(*
	One timed operation in a trace. Unlike a log record, a span has a lifecycle:
	  building - FB_Tracer owns it while the fluent chain fills it in,
	  running  - build hands it to the caller, who owns it while the work runs,
	  ended    - FB_Tracer.endSpan hands it to the provider for processing.
	The span owns every pointer member and releases them in free. A running span is read and
	changed only through FB_Tracer, such as getSpanContext, setSpanStatusOk and discardSpan,
	so callers never dereference it themselves. The methods left here belong to the tracing
	pipeline: the provider, samplers and processors.
*)
{attribute 'enable_dynamic_creation'}
FUNCTION_BLOCK FB_Span
VAR_INPUT
	// written by the tracer while the span is built
	name: POINTER TO FB_String;
	kind: E_SpanKind;
	startTimestamp: ULINT;
	endTimestamp: ULINT;
	traceId: POINTER TO FB_TraceId;
	spanId: POINTER TO FB_SpanId;
	traceState: POINTER TO FB_TraceState;

	// required if child span, must be omitted if root span
	parentSpanId: POINTER TO FB_SpanId;

	// describes the parent's remoteness, not this span's; see E_SpanFlags
	flags: UDINT;
	status: POINTER TO FB_Status;
END_VAR
VAR_OUTPUT
	attributes: FB_Attributes(maxCount := TcOtlp_GVL.DEFAULT_MAX_ATTRIBUTE_COUNT);
	links: FB_Links(maxCount := TcOtlp_GVL.DEFAULT_MAX_LINK_COUNT);
	resource: FB_Resource('');
	scope: FB_InstrumentationScope('', '', '');

	// span events have been deprecated, instead logs should be emitted with span context for correlation
	// events
	// droppedEventCount
END_VAR

(*
	Releases this span and clears the caller's pointer to it: call it as p^.delete(pSelf:=p).
	pSelf is cleared before the span is freed, so the caller never keeps a dangling pointer.
	A pointer to any other object is refused and left untouched, and nothing is released.
*)
METHOD delete : BOOL
VAR_IN_OUT
	pSelf: POINTER TO FB_Span;
END_VAR
VAR
	_pThis: POINTER TO FB_Span;
END_VAR
_pThis := THIS;
IF pSelf <> _pThis THEN
	RETURN;
END_IF

pSelf := 0;
__DELETE(_pThis);
delete := TRUE;
END_METHOD

//FB_Exit must be implemented explicitly. If there is an implementation, then the
//method is called before the controller removes the code of the function block instance
//(implicit call). The return value is not evaluated.
METHOD FB_Exit: BOOL
VAR_INPUT
    bInCopyCode: BOOL;  // TRUE: the exit method is called in order to leave the instance which will be copied afterwards (online change).
END_VAR
IF NOT bInCopyCode THEN
	THIS^.free();
END_IF
END_METHOD

(* Releases everything the span owns. Safe to call more than once. *)
METHOD free
IF THIS^.name <> 0 THEN THIS^.name^.delete(pSelf:=THIS^.name); END_IF
IF THIS^.traceId <> 0 THEN THIS^.traceId^.delete(pSelf:=THIS^.traceId); END_IF
IF THIS^.spanId <> 0 THEN THIS^.spanId^.delete(pSelf:=THIS^.spanId); END_IF
IF THIS^.traceState <> 0 THEN THIS^.traceState^.delete(pSelf:=THIS^.traceState); END_IF
IF THIS^.parentSpanId <> 0 THEN THIS^.parentSpanId^.delete(pSelf:=THIS^.parentSpanId); END_IF
IF THIS^.status <> 0 THEN THIS^.status^.delete(pSelf:=THIS^.status); END_IF
THIS^.attributes.free();
THIS^.links.free();
THIS^.scope.free();
THIS^.resource.free();
END_METHOD

(*
	Allocates a deep copy of this span, for a processor that keeps an ended span past onEnd.
	The copy owns copies of every member, so it stays valid after this span is released. This
	span is only read, apart from its links cursor. The caller owns pDest, which must be 0; on
	failure nothing is allocated and pDest is left alone.
*)
METHOD cloneTo : BOOL
VAR_IN_OUT
	pDest: POINTER TO FB_Span;
END_VAR
VAR_OUTPUT
	failureReason: E_SpanCloneFailureReason;
END_VAR
VAR
	_pClone: POINTER TO FB_Span;
	_pMessage: POINTER TO FB_String;
	_copied: BOOL;
	_attributesFailureReason: E_AttributesFailureReason;
	_linkFailureReason: E_LinkFailureReason;
END_VAR
cloneTo := FALSE;
failureReason := E_SpanCloneFailureReason.NA;

IF pDest <> 0 THEN
	failureReason := E_SpanCloneFailureReason.DESTINATION_ALREADY_ASSIGNED;
	RETURN;
END_IF

_pClone := __NEW(FB_Span);
IF _pClone = 0 THEN
	failureReason := E_SpanCloneFailureReason.MEMORY_ALLOCATION_FAILURE;
	RETURN;
END_IF

// the clone owns its members from here, so deleting it releases whatever was copied
_pClone^.kind := THIS^.kind;
_pClone^.startTimestamp := THIS^.startTimestamp;
_pClone^.endTimestamp := THIS^.endTimestamp;
_pClone^.flags := THIS^.flags;

_copied := (THIS^.name = 0 OR_ELSE ValueFactory.cloneString(
		pDest:=_pClone^.name,
		pSrc:=THIS^.name))
	AND_THEN (THIS^.traceId = 0 OR_ELSE ValueFactory.createTraceId(
		pDest:=_pClone^.traceId,
		pBytes:=ADR(THIS^.traceId^.bytes),
		nSize:=SIZEOF(THIS^.traceId^.bytes)))
	AND_THEN (THIS^.spanId = 0 OR_ELSE ValueFactory.createSpanId(
		pDest:=_pClone^.spanId,
		pBytes:=ADR(THIS^.spanId^.bytes),
		nSize:=SIZEOF(THIS^.spanId^.bytes)))
	AND_THEN (THIS^.parentSpanId = 0 OR_ELSE ValueFactory.createSpanId(
		pDest:=_pClone^.parentSpanId,
		pBytes:=ADR(THIS^.parentSpanId^.bytes),
		nSize:=SIZEOF(THIS^.parentSpanId^.bytes)))
	AND_THEN (THIS^.traceState = 0 OR_ELSE TraceStateFactory.clone(
		pDest:=_pClone^.traceState,
		pSrc:=THIS^.traceState))
	AND_THEN (THIS^.status = 0 OR_ELSE THIS^.status^.message = 0 OR_ELSE ValueFactory.cloneString(
		pDest:=_pMessage,
		pSrc:=THIS^.status^.message));
IF NOT _copied THEN
	IF _pMessage <> 0 THEN _pMessage^.delete(pSelf:=_pMessage); END_IF
	_pClone^.delete(pSelf:=_pClone);
	failureReason := E_SpanCloneFailureReason.VALUE_COPY_FAILURE;
	RETURN;
END_IF

IF THIS^.status <> 0 THEN
	_pClone^.status := __NEW(FB_Status(code:=THIS^.status^.code, message:=_pMessage));
	IF _pClone^.status = 0 THEN
		IF _pMessage <> 0 THEN _pMessage^.delete(pSelf:=_pMessage); END_IF
		_pClone^.delete(pSelf:=_pClone);
		failureReason := E_SpanCloneFailureReason.MEMORY_ALLOCATION_FAILURE;
		RETURN;
	END_IF
	_pMessage := 0;  // moved into the status
END_IF

IF NOT _pClone^.attributes.copyFrom(src:=THIS^.attributes, failureReason=>_attributesFailureReason) THEN
	_pClone^.delete(pSelf:=_pClone);
	IF _attributesFailureReason = E_AttributesFailureReason.MEMORY_ALLOCATION_FAILURE THEN
		failureReason := E_SpanCloneFailureReason.MEMORY_ALLOCATION_FAILURE;
	ELSE
		failureReason := E_SpanCloneFailureReason.ATTRIBUTE_COPY_FAILURE;
	END_IF
	RETURN;
END_IF

IF NOT _pClone^.links.copyFrom(src:=THIS^.links, failureReason=>_linkFailureReason) THEN
	_pClone^.delete(pSelf:=_pClone);
	IF _linkFailureReason = E_LinkFailureReason.MEMORY_ALLOCATION_FAILURE THEN
		failureReason := E_SpanCloneFailureReason.MEMORY_ALLOCATION_FAILURE;
	ELSE
		failureReason := E_SpanCloneFailureReason.LINK_COPY_FAILURE;
	END_IF
	RETURN;
END_IF

IF NOT _pClone^.resource.copyFrom(src:=THIS^.resource, failureResult=>_attributesFailureReason) THEN
	_pClone^.delete(pSelf:=_pClone);
	IF _attributesFailureReason = E_AttributesFailureReason.MEMORY_ALLOCATION_FAILURE THEN
		failureReason := E_SpanCloneFailureReason.MEMORY_ALLOCATION_FAILURE;
	ELSE
		failureReason := E_SpanCloneFailureReason.RESOURCE_COPY_FAILURE;
	END_IF
	RETURN;
END_IF

IF NOT _pClone^.scope.copyFrom(src:=THIS^.scope, failureResult=>_attributesFailureReason) THEN
	_pClone^.delete(pSelf:=_pClone);
	IF _attributesFailureReason = E_AttributesFailureReason.MEMORY_ALLOCATION_FAILURE THEN
		failureReason := E_SpanCloneFailureReason.MEMORY_ALLOCATION_FAILURE;
	ELSE
		failureReason := E_SpanCloneFailureReason.SCOPE_COPY_FAILURE;
	END_IF
	RETURN;
END_IF

// transfer ownership to the caller
pDest := _pClone;
_pClone := 0;
cloneTo := TRUE;
END_METHOD

(* TRUE when bit 0 of the trace flags, the W3C sampled flag, is set. *)
METHOD isSampled : BOOL
isSampled := (THIS^.flags AND 16#01) <> 0;
END_METHOD

(* Sets or clears bit 0 of the trace flags, the W3C sampled flag, and leaves the other bits. *)
METHOD setSampled
VAR_INPUT
	sampled: BOOL;
END_VAR
VAR CONSTANT
	TRACE_FLAG_SAMPLED: UDINT := 16#01;
END_VAR
IF sampled THEN
	THIS^.flags := THIS^.flags OR TRACE_FLAG_SAMPLED;
ELSE
	THIS^.flags := THIS^.flags AND NOT TRACE_FLAG_SAMPLED;
END_IF
END_METHOD

END_FUNCTION_BLOCK

(* stored: Version 1.1.0.1
   POU FB_Span: Id {17f1f0c3-d0bd-4cc5-82c0-c953a2faa69b}, SpecialFunc None
   Method delete: Id {6a97f055-36d8-4285-ad6e-08b9d3bfdaaf}
   Method FB_Exit: Id {fa780cfa-04fb-4c49-bd4c-b4e50dffd866}
   Method free: Id {8eaa02b8-df25-4adc-9c37-d019075ce71f}
   Method cloneTo: Id {8a52cd95-727f-4d26-979c-15f2ccdc0c38}
   Method isSampled: Id {c684c80b-3a08-4158-b7a3-910a9b9edce5}
   Method setSampled: Id {fefa0288-660b-4380-939e-fbe700e49687} *)
